(* IEC 61131-3 sources: PLC-IsaVODE/PLC-IsaVODE/samples/skeleton, 4 files *)

(* ---- 1-water_tank.st ---- *)
PROGRAM WTT
    VAR_INPUT
        x1, x2, f1, f2 : REAL;
    END_VAR
    VAR_OUTPUT
        V1, V2, P : BOOL;
    END_VAR

    IF (x1 >= H1) THEN
        V1 := 0;            (* Close inlet valve V1 if tank1 at high level *)
    ELSE
        IF (x1 <= L1) THEN
            V1 := 1;        (* Open V1 if tank1 at low level *)
        END_IF;
    END_IF;
    IF (x2 <= L2) THEN
        P := 1; V2 := 1;    (* If tank2 low, start pump P and open outlet valve V2 *)
    END_IF;
    IF (x1 <= LL OR f2 <= FL OR x2 >= H2) THEN
        P := 0; V2 := 0;    (* Emergency stop pump P and close V2 on underflow/overflow *)
    END_IF;
END_PROGRAM

(* ---- 2-for-and-while.st ---- *)
PROGRAM SimpleLoops
VAR
    i : INT;

    Sum1 : INT := 0;
    Sum2 : INT := 0;
    Sum3 : INT := 0;

    FirstBig : INT := 0;
    SkipSum : INT := 0;

    Count1 : INT := 0;
    Count2 : INT := 0;
    Count3 : INT := 0;

    x : INT := 0;
END_VAR

(* 1) Simple FOR *)
Sum1 := 0;
FOR i := 1 TO 5 DO
    Sum1 := Sum1 + i;
END_FOR;

(* 2) FOR with BY *)
Sum2 := 0;
FOR i := 1 TO 9 BY 2 DO
    Sum2 := Sum2 + i;
END_FOR;

(* 3) Reverse FOR *)
Sum3 := 0;
FOR i := 5 TO 1 BY -1 DO
    Sum3 := Sum3 + i;
END_FOR;

(* 4) FOR with EXIT *)
FirstBig := 0;
FOR i := 1 TO 10 DO
    IF i > 4 THEN
        FirstBig := i;
        EXIT;
    END_IF;
END_FOR;

(* 5) FOR with CONTINUE *)
SkipSum := 0;
FOR i := 1 TO 5 DO
    IF i = 3 THEN
        CONTINUE;
    END_IF;
    SkipSum := SkipSum + i;
END_FOR;

(* 6) Simple WHILE *)
x := 1;
Count1 := 0;
WHILE x <= 5 DO
    Count1 := Count1 + x;
    x := x + 1;
END_WHILE;

(* 7) WHILE with EXIT *)
x := 1;
Count2 := 0;
WHILE x <= 10 DO
    IF x > 4 THEN
        EXIT;
    END_IF;
    Count2 := Count2 + x;
    x := x + 1;
END_WHILE;

(* 8) WHILE with CONTINUE *)
x := 1;
Count3 := 0;
WHILE x <= 5 DO
    IF x = 3 THEN
        x := x + 1;
        CONTINUE;
    END_IF;
    Count3 := Count3 + x;
    x := x + 1;
END_WHILE;

END_PROGRAM

(* ---- 3-bohlender-artcile-reset-example.st ---- *)
PROGRAM RESET_BOHLENDER
	VAR RETAIN
	    fs : bool := true;
	END_VAR
	VAR
	    a : int := 0;
		b : int := 0;
	END_VAR

    IF fs THEN
    	b := 2;
    	fs := false;
    END_IF;
    a := 1234 / b;
END_PROGRAM

(* ---- 4-calibrate.st ---- *)
PROGRAM CALIBRATE
	VAR_INPUT
		X        : REAL;
		CO       : BOOL;
		CS       : BOOL;
		Y_OFFSET : REAL;
		Y_SCALE  : REAL;
	END_VAR

	VAR_OUTPUT
		Y 		 : REAL;
	END_VAR

	VAR RETAIN
		OFFSET   : REAL;
		SCALE    : REAL := 1.0;
	END_VAR

	IF CO THEN
		OFFSET := Y_OFFSET - X;
	ELSIF CS THEN
		SCALE := Y_SCALE / (X + OFFSET);
	END_IF;
	Y := (X + OFFSET) * SCALE;

END_PROGRAM
